TYPE T_ST_RJSEQ :
STRUCT
	ReadJobName:STRING;
	ReadLineNumber:WORD;
	ReadStepNumber:WORD;
END_STRUCT
END_TYPE

(* stored: Version 1.1.0.1, ProductVersion 3.1.4024.16
   DUT T_ST_RJSEQ: Id {219db4d2-6fb0-45a9-8ef4-a534ea714e62} *)
